(* IEC 61131-3 sources: kns-port-domestic/upstream/kns-pump-station/src/POUs/Station/FB_PumpProtection, 2 files *)

(* ---- FB_PumpProtection.decl.st ---- *)
// Назначение: защиты одного насоса (04 §10.3, 10.4): недогрузка по току («сухой ход насоса» —
//             работает на частоте не ниже rUnderloadSpeed_pct при токе ниже rUnderload_A дольше
//             tUnderload) с фиксацией до сброса насоса; перегрев обмотки — блокировка, пока сигнал
//             активен. Ток недостоверен — контроля нет; rUnderload_A = 0 — контроль выключен.
// Автор:      kr0nsch
// Версия:     0.1.0
// Документ:   docs/DESIGN.md, раздел 6.8; docs/04_algorithms.md, разделы 10.3, 10.4
FUNCTION_BLOCK FB_PumpProtection
VAR_INPUT
    xRunning      : BOOL;           // aitfPump[i].Running
    rSpeedAct_pct : REAL;           // aitfPump[i].SpeedAct
    rCurrent_A    : REAL;           // fbIT1n1.rValue_eu
    xCurrentValid : BOOL;           // fbIT1n1.xValid (нет связи — контроля нет)
    xOverheat     : BOOL;           // fbTS1n2.xValue
    xReset        : BOOL;           // импульс: GVL_Hmi.stP10nCmd.stCommon.xReset, HS501, xResetAll
    itfTime       : PL.I_TimeSource;
END_VAR
VAR_IN_OUT CONSTANT
    stCfg : ST_StationCfg;          // rUnderload_A (0 — выкл.), rUnderloadSpeed_pct, tUnderload
END_VAR
VAR_OUTPUT
    wInterlock       : WORD;        // KNS_ILK_UNDERLOAD (фиксация) OR KNS_ILK_OVERHEAT (пока сигнал)
    xUnderloadTrip   : BOOL;        // KNS1.ULn
    xUnderloadTiming : BOOL;
END_VAR
VAR
    fbUnderload : PL.FB_Delay;      // выдержка tUnderload
END_VAR
VAR_TEMP
    xCond : BOOL;                   // условие недогрузки до выдержки
END_VAR

(* ---- FB_PumpProtection.impl.st ---- *)
// 1. Сброс фиксации: импульс сброса насоса, кнопка HS501 или «Сбросить все» (04 §9.2). Насос под
//    блокировкой стоит, поэтому после сброса условие недогрузки отсчитывается заново
IF xReset THEN
    xUnderloadTrip := FALSE;
    fbUnderload.Preset(xValue := FALSE);
END_IF

// 2. Недогрузка (04 §10.3); неконечные ток и скорость — сравнения ложны, условия нет
xCond := stCfg.rUnderload_A > 0.0 AND xRunning AND xCurrentValid
         AND rSpeedAct_pct >= stCfg.rUnderloadSpeed_pct AND rCurrent_A < stCfg.rUnderload_A
         AND PL.F_IsFinite(rIn := rCurrent_A);
fbUnderload(xIn := xCond, tOnDelay := stCfg.tUnderload, itfTime := itfTime);
IF fbUnderload.xOut THEN
    xUnderloadTrip := TRUE;
END_IF
xUnderloadTiming := fbUnderload.xTimingOn;

// 3. Блокировки насоса: недогрузка — до сброса, перегрев — пока сигнал активен (04 §10.6)
wInterlock := 0;
IF xUnderloadTrip THEN
    wInterlock := wInterlock OR GVL_Const.KNS_ILK_UNDERLOAD;
END_IF
IF xOverheat THEN
    wInterlock := wInterlock OR GVL_Const.KNS_ILK_OVERHEAT;
END_IF
